{attribute 'qualified_only'}
//{attribute 'strict'}
{attribute 'to_string'}
TYPE E_CIP_DashStage_List :
(
	e00_NotSelected := 0,
	
	//CIP1
	e01_CIP1_Client_Drain_Product_Rest_Pipe,
	e02_CIP1_Client_Drain_Product_Rest_Sprinkler,
	
	//CIP2
	e03_CIP2_Local_Detergent_Fill,
	e04_CIP2_Local_Detergent_Condition,
	e05_CIP2_Client_Detergent_Fill,
	e06_CIP2_Client_Detergent_Condition_Pipe,	
	e07_CIP2_Client_Detergent_Condition_Sprinkler,	
	
	//CIP3
	e08_CIP3_Detergent_Collect,
	e09_CIP3_Detergent_Drain,
	e10_CIP3_Detergent_Clean_Pipe,
	e11_CIP3_Detergent_Clean_Sprinkler,
	
	//CIP4
	e12_CIP4_Local_DisInfection_Fill,
	e13_CIP4_Local_DisInfection_Condition,
	e14_CIP4_Client_DisInfection_Fill,
	e15_CIP4_Client_DisInfection_Condition_Pipe,	
	e16_CIP4_Client_DisInfection_Condition_Sprinkler,	
	
	//CIP5
	e17_CIP5_DisInfection_Collect,
	e18_CIP5_DisInfection_Drain,
	e19_CIP5_DisInfection_Clean_Pipe,
	e20_CIP5_DisInfection_Clean_Sprinkler,	
	
	
	eLast
);
END_TYPE

(* stored: Version 1.1.0.1, ProductVersion 3.1.4024.13
   DUT E_CIP_DashStage_List: Id {045304c0-0dd2-4309-8bac-7dc0272c5261} *)
